(* IEC 61131-3 sources: factorysim-public/codesys/acceptatie, 2 files *)

(* ---- IO.gvl.st ---- *)
(* Global Variable List "IO" — eigen werk, hoort bij de MVP-scène van FactorySim.
   Plak dit in een GVL met de naam IO. De volgorde en namen komen overeen met
   src/FactorySim.App/tagmap.json. *)
VAR_GLOBAL
    (* App -> PLC: Coils 0..7 van het Modbus TCP Slave Device *)
    iStart       : BOOL;    (* Coil 0: startknop (puls) *)
    iStop        : BOOL;    (* Coil 1: stopknop, TRUE = ingedrukt *)
    iAtPusher    : BOOL;    (* Coil 2: photo-eye, doos voor de pusher *)
    iHighBox     : BOOL;    (* Coil 3: hoge photo-eye, doos is hoog *)
    iPusherBack  : BOOL;    (* Coil 4: pusher ingetrokken *)
    iPusherFront : BOOL;    (* Coil 5: pusher uitgeschoven *)
    iSimRunning  : BOOL;    (* Coil 6: simulatie draait *)
    iSpare       : BOOL;    (* Coil 7: reserve *)

    (* PLC -> App: Discrete Inputs 0..7 van het Modbus TCP Slave Device *)
    oConveyor    : BOOL;    (* Discrete Input 0: band aan *)
    oPusher      : BOOL;    (* Discrete Input 1: pusher uitschuiven *)
    oEmitter     : BOOL;    (* Discrete Input 2: dozen spawnen *)
    oRunLamp     : BOOL;    (* Discrete Input 3: lamp in bedrijf *)
    oSpare1      : BOOL;
    oSpare2      : BOOL;
    oSpare3      : BOOL;
    oSpare4      : BOOL;
END_VAR

(* ---- PLC_PRG.st ---- *)
(* Acceptatieprogramma voor de MVP-scène van FactorySim — eigen werk.
   Start/stop en sorteren op hoogte: hoge dozen gaan via de pusher naar de zijbaan,
   lage dozen rijden door. Dezelfde logica zit in tools/fake_plc/fake_plc.py (modus sorter).

   In CODESYS: het declaratiedeel hieronder in het bovenste venster van PLC_PRG plakken,
   het programmadeel in het onderste. *)

(* ---------- Declaratie ---------- *)
PROGRAM PLC_PRG
VAR
    bRun    : BOOL;         (* installatie in bedrijf *)
    nStep   : INT := 0;     (* 0 = transport, 10 = duwen, 20 = terug *)
    tonPush : TON;          (* bewaking: pusher haalt zijn eindstand niet *)
    bFault  : BOOL;
    nSorted : UDINT;        (* aantal uitgesorteerde dozen *)
END_VAR

(* ---------- Programma ---------- *)

(* Start/stop: stop dominant, alleen als de simulatie draait *)
IF IO.iStop OR NOT IO.iSimRunning OR bFault THEN
    bRun := FALSE;
ELSIF IO.iStart THEN
    bRun := TRUE;
END_IF

(* Fout resetten met Start terwijl Stop is losgelaten *)
IF bFault AND IO.iStart AND NOT IO.iStop THEN
    bFault := FALSE;
    nStep  := 0;
END_IF

(* Sorteerstap *)
CASE nStep OF
    0:  (* transport *)
        IF bRun AND IO.iAtPusher AND IO.iHighBox AND IO.iPusherBack THEN
            nStep := 10;
        END_IF

    10: (* band stil, pusher uit *)
        IF IO.iPusherFront THEN
            nSorted := nSorted + 1;
            nStep := 20;
        END_IF

    20: (* pusher terug *)
        IF IO.iPusherBack THEN
            nStep := 0;
        END_IF
END_CASE

(* Bewaking: de pusher moet binnen 3 s zijn eindstand halen.
   Alleen terwijl de simulatie draait, zodat pauzeren geen fout geeft. *)
tonPush(IN := ((nStep = 10) OR (nStep = 20)) AND IO.iSimRunning, PT := T#3S);
IF tonPush.Q THEN
    bFault := TRUE;
    nStep  := 0;
END_IF

(* Uitgangen *)
IO.oConveyor := bRun AND (nStep = 0);
IO.oPusher   := (nStep = 10);
IO.oEmitter  := bRun;
IO.oRunLamp  := bRun;
